TYPE ST_Command :
STRUCT
	bEnable: BOOL;
	bExecute: BOOL;
	bContinuousupdate: BOOL;
END_STRUCT
END_TYPE

(* stored: Version 1.1.0.1, ProductVersion 3.1.4024.12
   DUT ST_Command: Id {1dfcc98d-ec82-4c48-87be-d61db0310a67} *)
